Staubli VAL3: HMI_progEdit.dtx

mdesc mNomSpeed
string sSelProg
bool bBack
public bool bBool[9]
public bool bInsert[16]
num nPageIndex
num nPageNum
public num nLstValue
string sLstValue
string sList
bool bToSave
string sPageNum
string sPageIndex
public bool bTRAJ[7]
string sPgIndexTRAJ
string sPageTRAJ
num nPgIndexTRAJ
num nPgNumTRAJ
string sTRAJList
string sInsertItem
string sPgIndexPROG
string sPagePROG
num nPgIndexPROG
num nPgNumPROG
string sPROGList
string sIFType[3]
public num nIFValue[3]
string sIFIndex[3]
string sANDOR1
string sANDOR2
bool bIFConfirm
bool bIFCancel
string sLastANDOR2
string sLastANDOR1
bool bSwitchOK
bool bSwitchCancel
string sIOList
string sSwitchValue
num nCaseValue
num nFORValue
string sForValue
bool bSelProg
bool bSelTraj
bool bBindTRAJ
bool bBindProg
num nSelType
